// TIA Portal V20 export
Screen "RobotService_Zone04"  1276x673
  ScreenItem "Line_Header_X0_Y64" at 0,64 size 1280x0  Type=HmiLine
  ScreenItem "permanentareaborderrectangle" at 0,0 size 0x0  Type=HmiRectangle
  ScreenItem "Button_Back" at 2,2 size 90x60  Type=HmiButton
  ScreenItem "Title_ScreenOverview_X390_Y2_3" at 375,5 size 510x57  Type=HmiTextBox
  ScreenItem "Faceplate container_2" at 1128,69 size 127x580  Type=HmiFaceplateContainer
  ScreenItem "130RB02" at 314,69 size 193x297  Type=HmiFaceplateContainer
  ScreenItem "130RB01" at 28,69 size 193x297  Type=HmiFaceplateContainer
  ScreenItem "140RB01" at 601,69 size 193x297  Type=HmiFaceplateContainer
